SUBAPPLICATION Name
  (* Standard: 61499-1; Description: Copyright (c) 2026 Martin Erich Jobst This program and the accompanying materials are made available under the terms of the Eclipse Public License 2.0 which is available at https://www.eclipse.org/legal/epl-2.0/ SPDX-License-Identifier: EPL-2.0 *)
  (* Version 1.0, 2026-11-18, Martin Jobst *)
  PACKAGE lib::VarConfigInstance;
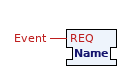
  EVENT_INPUT
    REQ;
  END_EVENT
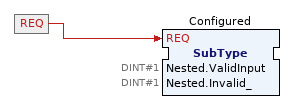
  SUBAPPS
    Configured : lib::VarConfigInstance::support::SubType(Nested.ValidInput := DINT#1, Nested.Invalid_ := DINT#1);
  END_SUBAPPS
  EVENT_CONNECTIONS
    REQ TO Configured.REQ;
  END_CONNECTIONS
END_SUBAPPLICATION
